FUNCTION F_ModuloDistance : DINT
(*
Function for calculate modulo distance.

Constructor: 	Patryk Panylo
Company:		E. Riexinger GmbH
Date:			20.01.2014
Version:		1.00

Date:			Revision:		Who:				Comment
dd.mm.yyyy		x.xx			Initials			comment

*)

VAR_INPUT
	dwCurrentValue			:DWORD;
	dwOldValue				:DWORD;
	dwModuloValue			:DWORD;
END_VAR
VAR
	dwPosDistance			:DWORD;

END_VAR


F_ModuloDistance := DWORD_TO_DINT(dwCurrentValue - dwOldValue);

IF dwModuloValue <> 0
THEN
	dwPosDistance := F_ModDW(dwCurrentValue - dwOldValue, dwModuloValue);
	
	F_ModuloDistance := DWORD_TO_DINT(dwPosDistance);
	
	IF dwPosDistance > (dwModuloValue / 2) 
	THEN
		F_ModuloDistance := -DWORD_TO_DINT(dwModuloValue - dwPosDistance);
	END_IF
	
END_IF

END_FUNCTION

(* stored: Version 1.1.0.1, ProductVersion 3.1.4024.15
   POU F_ModuloDistance: Id {2d673631-b9c3-49a6-98e3-98ae42a359ba}, SpecialFunc None *)
